(* IEC 61131-3 sources: model-first-plc-agent-ai/results/T2-W-10, 2 files *)

(* ---- a1_code.st ---- *)
FUNCTION_BLOCK FillingRuntime
VAR_INPUT
    start : BOOL;
    stop : BOOL;
    LSH : BOOL;
    LSHH : BOOL;
    TimerDuration : TIME;
END_VAR
VAR_OUTPUT
    fill_valve : BOOL;
    discharge_valve : BOOL;
END_VAR
VAR
    x0 : BOOL := TRUE;
    x1 : BOOL := FALSE;
    t1 : BOOL;
    t2 : BOOL;
    timer_done : BOOL := FALSE;
    FillingTimer : TON;
END_VAR

(* Evaluate the start transition from the current situation. *)
t1 := x0 AND start AND NOT stop AND NOT LSHH;

(* Begin timing in the same scan that the filling step is entered. *)
FillingTimer(IN := x1 OR t1, PT := TimerDuration);

(* The owned condition is FALSE at the instant x1 becomes active. *)
timer_done := x1 AND FillingTimer.Q;

t2 := x1 AND (stop OR LSHH OR timer_done);

(* Apply transitions using the preceding situation. *)
IF t2 THEN
    x0 := TRUE;
    x1 := FALSE;
ELSIF t1 THEN
    x0 := FALSE;
    x1 := TRUE;
END_IF;

(* Reset the timer immediately whenever its owning step is inactive. *)
IF NOT x1 THEN
    FillingTimer(IN := FALSE, PT := TimerDuration);
    timer_done := FALSE;
END_IF;

fill_valve := x1;
discharge_valve := FALSE;

END_FUNCTION_BLOCK

PROGRAM Main
VAR
    StartCommand AT %IX100.0 : BOOL;
    StopCommand AT %IX100.1 : BOOL;
    LSH AT %IX100.2 : BOOL;
    LSHH AT %IX100.3 : BOOL;
    FillValve AT %QX100.0 : BOOL;
    DischargeValve AT %QX100.1 : BOOL;
END_VAR
VAR
    (* Configurable filling-duration parameter. *)
    TimerDuration : TIME := T#5s;
    StartEdge : R_TRIG;
    Controller : FillingRuntime;
END_VAR

StartEdge(CLK := StartCommand);

Controller(
    start := StartEdge.Q,
    stop := StopCommand,
    LSH := LSH,
    LSHH := LSHH,
    TimerDuration := TimerDuration
);

FillValve := Controller.fill_valve;
DischargeValve := Controller.discharge_valve;

END_PROGRAM

(* ---- a2_code.st ---- *)
FUNCTION_BLOCK FB_TimedTankFilling
VAR_INPUT
    StartCommand : BOOL;
    StopCommand : BOOL;
    LSH : BOOL;
    LSHH : BOOL;
    TimerDuration : TIME;
END_VAR
VAR_OUTPUT
    fill_valve : BOOL;
    discharge_valve : BOOL;
END_VAR
VAR
    StartEdge : R_TRIG;
    FillTimer : TON;
    start : BOOL;
    stop : BOOL;
    timer_done : BOOL;
    CurrentState : INT := 0;
END_VAR

StartEdge(CLK := StartCommand);
start := StartEdge.Q;
stop := StopCommand;

IF stop THEN
    CurrentState := 0;
ELSE
    CASE CurrentState OF
        0:
            IF start AND NOT LSHH THEN
                CurrentState := 1;
            END_IF;

        1:
            IF LSHH THEN
                CurrentState := 0;
            END_IF;

        ELSE
            CurrentState := 0;
    END_CASE;
END_IF;

FillTimer(IN := (CurrentState = 1), PT := TimerDuration);
timer_done := FillTimer.Q;

IF (CurrentState = 1) AND timer_done THEN
    CurrentState := 0;
END_IF;

IF CurrentState = 0 THEN
    FillTimer(IN := FALSE, PT := TimerDuration);
    timer_done := FALSE;
END_IF;

fill_valve := (CurrentState = 1);
discharge_valve := FALSE;

END_FUNCTION_BLOCK

PROGRAM Main
VAR
    StartCommand AT %IX100.0 : BOOL;
    StopCommand AT %IX100.1 : BOOL;
    LSH AT %IX100.2 : BOOL;
    LSHH AT %IX100.3 : BOOL;
    FillValve AT %QX100.0 : BOOL;
    DischargeValve AT %QX100.1 : BOOL;
END_VAR
VAR
    TimerDuration : TIME := T#10s;
    TankController : FB_TimedTankFilling;
END_VAR

TankController(
    StartCommand := StartCommand,
    StopCommand := StopCommand,
    LSH := LSH,
    LSHH := LSHH,
    TimerDuration := TimerDuration
);

FillValve := TankController.fill_valve;
DischargeValve := TankController.discharge_valve;

END_PROGRAM
